{attribute 'qualified_only'}
VAR_GLOBAL CONSTANT
	rTime2Seconds	:	REAL	:=	0.001;
	rSeconds2Time	:	REAL	:=	1000;
END_VAR

(* stored: Version 1.1.0.1, ProductVersion 3.1.4024.9
   GVL CONVERSIONS: Id {11182d4b-a82b-4df1-a41f-27597d1f24fd} *)
